{attribute 'qualified_only'}
{attribute 'strict'}
{attribute 'to_string'}
TYPE E_Element_Type :
(
eNotSelected := 0,
eTank,
eTriBlender,
eLine
);
END_TYPE

(* stored: Version 1.1.0.1, ProductVersion 3.1.4024.12
   DUT E_Element_Type: Id {5c898ead-6018-47b3-bcc4-52428c4260bb} *)
